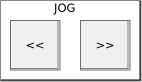
VISUALIZATION JOG  // 142x82
    Rectangle (-10,0 150x80), "JOG"
    Button (10,20 50x50), "<<"
        tap MAIN.Track.Jog.JogBackwards
    Button (80,20 50x50), ">>"
        tap MAIN.Track.Jog.JogForward
END_VISUALIZATION

(* stored: Version 1.1.0.1, ProductVersion 3.1.4024.16
   Visu JOG: Id {a42888f2-16bf-4ead-90e0-d7fdf305564d} *)
